Fanuc KAREL source: kd00023.compact.KL

PROGRAM KD00023
%STACKSIZE=65535
%PRIORITY=65535
%NOLOCKGROUP
VAR
I : INTEGER
J : INTEGER
B : BOOLEAN
R : REAL
S : STRING[80]
SAVED : INTEGER
BEGIN
I=SAVED
END KD00023
